(* IEC 61131-3 sources: volt/packages/volt-lsp-iec/test-corpus/pro2193/Device/Plc Logic/Application/09 Misc/Library Manager/L_TT1P_TechnologyModules (part 6) *)

(* ---- L_TT1P_WINDERTENSIONCTRLHIGH.pou ---- *)
FUNCTION_BLOCK L_TT1P_WINDERTENSIONCTRLHIGH EXTENDS TM_Winder
VAR_INPUT
	XENABLEINTERNALCONTROL : BOOL;
	XENABLE : BOOL;
	SCCTRLABC : scCtrl_ABC;
	XRESETERROR : BOOL;
	XREGULATORON : BOOL;
	XSTOP : BOOL;
	XHALT : BOOL;
	SCPAR : L_TT1P_scPar_WinderTensionCtrlHigh;
	MATERIALCOUNTERAXIS : L_MC1P_IAXIS_REF_POOL;
	SCACCESSPOINTS : L_TT1P_scAP_WinderTensionCtrlHigh;
	XMATERIALFEEDING : BOOL;
	XWINDINGDIRECTION : BOOL;
	XWINDINGDIRECTIONSTANDSTILL : BOOL;
	XLOADDIAM : BOOL;
	LRSETDIAM : LREAL;
	XHOLDDIAM : BOOL;
	XDIAMCALCREDUCED : BOOL;
	XSETMATERIALCOUNTER : BOOL;
	XWEBBREAKMONIT : BOOL;
	XJOGLINEPOS : BOOL;
	XJOGLINENEG : BOOL;
	XTRIMLINEPOS : BOOL;
	XTRIMLINENEG : BOOL;
	XSYNCLINEVEL : BOOL;
	XTENSCURVE : BOOL;
	LRSETTENS : LREAL;
	LRSETLINEVEL : LREAL;
	XTENSCTRL : BOOL;
	XFRICCMPS : BOOL;
	XACCCMPS : BOOL;
	LRMINERTIAADAPT : LREAL;
	LRACTTENSIN : LREAL;
	LRSETFRICADAPT : LREAL;
	LRTENSCTRLINFLUENCE : LREAL;
	XRESETPICTRL : BOOL;
	XRESETICTRL : BOOL;
	XEXECUTEIDENTFRIC : BOOL;
	XEXECUTEIDENTMINERTIA : BOOL;
	XADAPTSPDCTRLGAIN : BOOL;
	LRADAPTSPDCTRLGAINFACTOR : LREAL := 1;
END_VAR
VAR_OUTPUT
	XINTERNALCONTROLACTIVE : BOOL;
	ETMSTATE : L_TT1P_States;
	SCSTATUSABC : scStatus_ABC;
	XERROR : BOOL;
	XWARNING : BOOL;
	EERRORID : L_IE1P_Error;
	SCERRORINFO : L_TT1P_scErrorInfo;
	XAXISENABLED : BOOL;
	SCSIGNALFLOW : L_TT1P_scSF_WinderTensionCtrlHigh;
	XDONE : BOOL;
	XBUSY : BOOL;
	XSYNCHRONISED : BOOL;
	XACCDECSYNC : BOOL;
	XUNWIND : BOOL;
	XWEBBREAK : BOOL;
	XHOLDDIAMACTIVE : BOOL;
	XDIAMMAX : BOOL;
	XDIAMMIN : BOOL;
	LRSETDIAMOUT : LREAL;
	LRSETDIAMSCALEDOUT : LREAL;
	LRMATERIALCOUNTER : LREAL;
	LRSETLINEVELSCALEDOUT : LREAL;
	LRACTTOTALTRQSCALED : LREAL;
	LRWNDSPDREF : LREAL;
	XWNDSPDLIMIT : BOOL;
	LRLIMITLINEVEL : LREAL;
	LRSETMINERTIAOUT : LREAL;
	LRSETTENSSCALEDOUT : LREAL;
	LRSETTENSTRQSCALEDOUT : LREAL;
	LRSETFRICTRQSCALEDOUT : LREAL;
	LRSETACCTRQSCALEDOUT : LREAL;
	LRACTTENSSCALED : LREAL;
	LRSETTENSCTRLSCALEDOUT : LREAL;
	LRIDENTMINERTIA : LREAL;
	LRSETSPDCTRLGAINADAPTOUT : LREAL;
END_VAR
VAR_IN_OUT
	AXIS : AXIS_REF;
	PERSISTENTVAR : L_TT1P_PersistentVarWinder;
	ALRFRICTIONCURVE1 : ARRAY [1..66] OF LREAL;
	ALRFRICTIONCURVE2 : ARRAY [1..66] OF LREAL;
	ALRFRICTIONCURVE3 : ARRAY [1..66] OF LREAL;
	ALRFRICTIONCURVE4 : ARRAY [1..66] OF LREAL;
END_VAR
VAR
	TM_INT : _TM_WinderTensionCtrlHigh;
	PPAR : POINTER TO L_TT1P_scPar_WinderTensionCtrlHigh;
	PPAR_INT : POINTER TO L_TT1P_scPar_WinderTensionCtrlHigh;
	XISHOMED : BOOL;
	XHOMEEXECUTE : BOOL;
	XHOMEABSSWITCH : BOOL;
	XJOGPOS : BOOL;
	XJOGNEG : BOOL;
END_VAR
END_FUNCTION_BLOCK

METHOD CALL_COUPLINGREELSPEEDLIMIT
END_METHOD

METHOD CALL_DECOUPLINGREELSPEEDLIMIT
END_METHOD

METHOD GET_ESTATE : L_TT1P_States
END_METHOD

METHOD GET_ETMSTATE : L_TT1P_States
END_METHOD

METHOD GET_LRACTACCTRQ : LREAL
END_METHOD

METHOD GET_LRACTFRICTRQ : LREAL
END_METHOD

METHOD GET_LRACTMOTORTORQUE : LREAL
END_METHOD

METHOD GET_LRACTTENSTRQ : LREAL
END_METHOD

METHOD GET_LRCALCDIAMDIST : LREAL
END_METHOD

METHOD GET_LRCALCDIAMLINESPEED : LREAL
END_METHOD

METHOD GET_LRCALCDIAMREELSPEED : LREAL
END_METHOD

METHOD GET_LRFEEDCONSTANT : LREAL
END_METHOD

METHOD GET_LRLOWERSPEEDLIMIT : LREAL
END_METHOD

METHOD GET_LRMOTORTORQUEREF : LREAL
END_METHOD

METHOD GET_LRRAMPGENOUT : LREAL
END_METHOD

METHOD GET_LRREELSPEEDREF : LREAL
END_METHOD

METHOD GET_LRSETMOTORTORQUE : LREAL
END_METHOD

METHOD GET_LRSETSPEEDCTRLGAINADAPT : LREAL
END_METHOD

METHOD GET_LRSETTOTALTORQUE : LREAL
END_METHOD

METHOD GET_LRSPEEDLOWERLIMIT : LREAL
END_METHOD

METHOD GET_LRSPEEDUPPERLIMIT : LREAL
END_METHOD

METHOD GET_LRTASKCYCLE : LREAL
END_METHOD

METHOD GET_LRTENSCTRLOUT : LREAL
END_METHOD

METHOD GET_LRTENSCURVEOUT : LREAL
END_METHOD

METHOD GET_LRUPPERSPEEDLIMIT : LREAL
END_METHOD

METHOD GET_LRVARMINERTIASCALED : LREAL
END_METHOD

METHOD GET_LRWINDERTORQUEREF : LREAL
END_METHOD

METHOD GET_XCOMMUNICATION : BOOL
END_METHOD

METHOD GET_XDIAMWEBBREAKENABLE : BOOL
VAR_OUTPUT
	XUNIDIRECT : BOOL;
	XUNWINDACTIVE : BOOL;
END_VAR
END_METHOD

METHOD RESET_SYSTEMFAULT
END_METHOD

METHOD SET_SYSTEMFAULT
VAR_INPUT
	IN : L_IE1P_Error;
END_VAR
END_METHOD

METHOD SET_ALRPROCESSCTRLXVALUES
VAR_INPUT
	ALRPROCESSCTRLXVALUES : ARRAY [1..5] OF LREAL := [5(0)];
END_VAR
END_METHOD

METHOD SET_ALRPROCESSCTRLYVALUES
VAR_INPUT
	ALRPROCESSCTRLYVALUES : ARRAY [1..5] OF LREAL := [1, 4(0)];
END_VAR
END_METHOD

METHOD SET_ESTATE
VAR_INPUT
	IN : L_TT1P_States;
END_VAR
END_METHOD

METHOD SET_LRFEEDCONSTANT
VAR_INPUT
	LRIN : LREAL := 0;
END_VAR
END_METHOD

METHOD SET_LRPICTRLINTVALUE
VAR_INPUT
	LRIN : LREAL := 0;
END_VAR
END_METHOD

METHOD SET_LRPROCESSCTRLACC
VAR_INPUT
	LRPROCESSCTRLACC : LREAL := 0.0;
END_VAR
END_METHOD

METHOD SET_LRPROCESSCTRLDEC
VAR_INPUT
	LRPROCESSCTRLDEC : LREAL := 0.0;
END_VAR
END_METHOD

METHOD SET_LRPROCESSCTRLGAINADAPT
VAR_INPUT
	LRPROCESSCTRLGAINADAPT : LREAL := 1;
END_VAR
END_METHOD

METHOD SET_LRPROCESSCTRLINTVALUE
VAR_INPUT
	LRPROCESSCTRLINTVALUE : LREAL := 0.0;
END_VAR
END_METHOD

METHOD SET_LRPROCESSCTRLREDGAIN
VAR_INPUT
	LRPROCESSCTRLREDGAIN : LREAL := 0.0;
END_VAR
END_METHOD

METHOD SET_LRPROCESSCTRLREDRANGE
VAR_INPUT
	LRPROCESSCTRLREDRANGE : LREAL := 0.0;
END_VAR
END_METHOD

METHOD SET_LRREFERENCEMOTORTORQUE
VAR_INPUT
	LRIN : LREAL := 0;
END_VAR
END_METHOD

METHOD SET_LRREFERENCEREELSPEED
VAR_INPUT
	LRIN : LREAL := 0;
END_VAR
END_METHOD

METHOD SET_LRSPEEDOFFSET
VAR_INPUT
	LRIN : LREAL := 0;
END_VAR
END_METHOD

METHOD SET_LRTORQUEOFFSET
VAR_INPUT
	LRIN : LREAL := 0;
END_VAR
END_METHOD

METHOD SET_RPROCESSCTRLDELAYTIME
VAR_INPUT
	RPROCESSCTRLDELAYTIME : REAL := 0.0;
END_VAR
END_METHOD

METHOD SET_RPROCESSCTRLRATEDTIME
VAR_INPUT
	RPROCESSCTRLRATEDTIME : REAL := 0.0;
END_VAR
END_METHOD

METHOD SET_XPICTRLLOADINTVALUE
VAR_INPUT
	XIN : BOOL := FALSE;
END_VAR
END_METHOD

METHOD SET_XPROCESSCTRLLOADINTVALUE
VAR_INPUT
	XPROCESSCTRLLOADINTVALUE : BOOL := FALSE;
END_VAR
END_METHOD

METHOD SET_XSPEEDLIMITENABLEDEXT
VAR_INPUT
	XIN : BOOL := TRUE;
END_VAR
END_METHOD

METHOD SET_XWEBBREAK
VAR_INPUT
	XIN : BOOL := FALSE;
END_VAR
END_METHOD

(* ---- L_TT1P_WINDERTENSIONCTRLSTATE.pou ---- *)
FUNCTION_BLOCK L_TT1P_WINDERTENSIONCTRLSTATE EXTENDS TM_Winder
VAR_INPUT
	XENABLEINTERNALCONTROL : BOOL;
	XENABLE : BOOL;
	SCCTRLABC : scCtrl_ABC;
	XRESETERROR : BOOL;
	XREGULATORON : BOOL;
	XSTOP : BOOL;
	XHALT : BOOL;
	SCPAR : L_TT1P_scPar_WinderTensionCtrlState;
	MATERIALCOUNTERAXIS : L_MC1P_IAXIS_REF_POOL;
	SCACCESSPOINTS : L_TT1P_scAP_WinderTensionCtrlState;
	XMATERIALFEEDING : BOOL;
	XWINDINGDIRECTION : BOOL;
	XWINDINGDIRECTIONSTANDSTILL : BOOL;
	XLOADDIAM : BOOL;
	LRSETDIAM : LREAL;
	XHOLDDIAM : BOOL;
	XDIAMCALCREDUCED : BOOL;
	XSETMATERIALCOUNTER : BOOL;
	XWEBBREAKMONIT : BOOL;
	XJOGLINEPOS : BOOL;
	XJOGLINENEG : BOOL;
	XTRIMLINEPOS : BOOL;
	XTRIMLINENEG : BOOL;
	XSYNCLINEVEL : BOOL;
	XTENSCURVE : BOOL;
	LRSETTENS : LREAL;
	LRSETLINEVEL : LREAL;
	XTENSCTRL : BOOL;
	XFRICCMPS : BOOL;
	XACCCMPS : BOOL;
	LRMINERTIAADAPT : LREAL := 1;
	LRACTTENSIN : LREAL;
	LRSETFRICADAPT : LREAL;
	LRTENSCTRLINFLUENCE : LREAL;
	XRESETPICTRL : BOOL;
	XRESETICTRL : BOOL;
	XEXECUTEIDENTFRIC : BOOL;
END_VAR
VAR_OUTPUT
	XINTERNALCONTROLACTIVE : BOOL;
	ETMSTATE : L_TT1P_States;
	SCSTATUSABC : scStatus_ABC;
	XERROR : BOOL;
	XWARNING : BOOL;
	EERRORID : L_IE1P_Error;
	SCERRORINFO : L_TT1P_scErrorInfo;
	XAXISENABLED : BOOL;
	SCSIGNALFLOW : L_TT1P_scSF_WinderTensionCtrlState;
	XDONE : BOOL;
	XBUSY : BOOL;
	XSYNCHRONISED : BOOL;
	XACCDECSYNC : BOOL;
	XUNWIND : BOOL;
	XWEBBREAK : BOOL;
	XHOLDDIAMACTIVE : BOOL;
	XDIAMMAX : BOOL;
	XDIAMMIN : BOOL;
	LRSETDIAMOUT : LREAL;
	LRSETDIAMSCALEDOUT : LREAL;
	LRMATERIALCOUNTER : LREAL;
	LRSETLINEVELSCALEDOUT : LREAL;
	LRACTTOTALTRQSCALED : LREAL;
	LRWNDSPDREF : LREAL;
	XWNDSPDLIMIT : BOOL;
	LRLIMITLINEVEL : LREAL;
	LRSETMINERTIAOUT : LREAL;
	LRSETTENSSCALEDOUT : LREAL;
	LRSETTENSTRQSCALEDOUT : LREAL;
	LRSETFRICTRQSCALEDOUT : LREAL;
	LRSETACCTRQSCALEDOUT : LREAL;
	LRACTTENSSCALED : LREAL;
	LRSETTENSCTRLSCALEDOUT : LREAL;
END_VAR
VAR_IN_OUT
	AXIS : AXIS_REF;
	PERSISTENTVAR : L_TT1P_PersistentVarWinder;
	ALRFRICTIONCURVE1 : ARRAY [1..66] OF LREAL;
	ALRFRICTIONCURVE2 : ARRAY [1..66] OF LREAL;
	ALRFRICTIONCURVE3 : ARRAY [1..66] OF LREAL;
	ALRFRICTIONCURVE4 : ARRAY [1..66] OF LREAL;
END_VAR
VAR
	TM_INT : _TM_WinderTensionCtrlState;
	PPAR : POINTER TO L_TT1P_scPar_WinderTensionCtrlState;
	PPAR_INT : POINTER TO L_TT1P_scPar_WinderTensionCtrlState;
	XISHOMED : BOOL;
	XHOMEEXECUTE : BOOL;
	XHOMEABSSWITCH : BOOL;
	XJOGPOS : BOOL;
	XJOGNEG : BOOL;
END_VAR
END_FUNCTION_BLOCK

METHOD CALL_COUPLINGREELSPEEDLIMIT
END_METHOD

METHOD CALL_DECOUPLINGREELSPEEDLIMIT
END_METHOD

METHOD GET_ESTATE : L_TT1P_States
END_METHOD

METHOD GET_ETMSTATE : L_TT1P_States
END_METHOD

METHOD GET_LRACTACCTRQ : LREAL
END_METHOD

METHOD GET_LRACTFRICTRQ : LREAL
END_METHOD

METHOD GET_LRACTMOTORTORQUE : LREAL
END_METHOD

METHOD GET_LRACTTENSTRQ : LREAL
END_METHOD

METHOD GET_LRCALCDIAMDIST : LREAL
END_METHOD

METHOD GET_LRCALCDIAMLINESPEED : LREAL
END_METHOD

METHOD GET_LRCALCDIAMREELSPEED : LREAL
END_METHOD

METHOD GET_LRFEEDCONSTANT : LREAL
END_METHOD

METHOD GET_LRLOWERSPEEDLIMIT : LREAL
END_METHOD

METHOD GET_LRMOTORTORQUEREF : LREAL
END_METHOD

METHOD GET_LRRAMPGENOUT : LREAL
END_METHOD

METHOD GET_LRREELSPEEDREF : LREAL
END_METHOD

METHOD GET_LRSETMOTORTORQUE : LREAL
END_METHOD

METHOD GET_LRSETSPEEDCTRLGAINADAPT : LREAL
END_METHOD

METHOD GET_LRSETTOTALTORQUE : LREAL
END_METHOD

METHOD GET_LRSPEEDLOWERLIMIT : LREAL
END_METHOD

METHOD GET_LRSPEEDUPPERLIMIT : LREAL
END_METHOD

METHOD GET_LRTASKCYCLE : LREAL
END_METHOD

METHOD GET_LRTENSCTRLOUT : LREAL
END_METHOD

METHOD GET_LRTENSCURVEOUT : LREAL
END_METHOD

METHOD GET_LRUPPERSPEEDLIMIT : LREAL
END_METHOD

METHOD GET_LRVARMINERTIASCALED : LREAL
END_METHOD

METHOD GET_LRWINDERTORQUEREF : LREAL
END_METHOD

METHOD GET_XCOMMUNICATION : BOOL
END_METHOD

METHOD GET_XDIAMWEBBREAKENABLE : BOOL
VAR_OUTPUT
	XUNIDIRECT : BOOL;
	XUNWINDACTIVE : BOOL;
END_VAR
END_METHOD

METHOD RESET_SYSTEMFAULT
END_METHOD

METHOD SET_SYSTEMFAULT
VAR_INPUT
	IN : L_IE1P_Error;
END_VAR
END_METHOD

METHOD SET_ALRPROCESSCTRLXVALUES
VAR_INPUT
	ALRPROCESSCTRLXVALUES : ARRAY [1..5] OF LREAL := [5(0)];
END_VAR
END_METHOD

METHOD SET_ALRPROCESSCTRLYVALUES
VAR_INPUT
	ALRPROCESSCTRLYVALUES : ARRAY [1..5] OF LREAL := [1, 4(0)];
END_VAR
END_METHOD

METHOD SET_ESTATE
VAR_INPUT
	IN : L_TT1P_States;
END_VAR
END_METHOD

METHOD SET_LRFEEDCONSTANT
VAR_INPUT
	LRIN : LREAL := 0;
END_VAR
END_METHOD

METHOD SET_LRPICTRLINTVALUE
VAR_INPUT
	LRIN : LREAL := 0;
END_VAR
END_METHOD

METHOD SET_LRPROCESSCTRLACC
VAR_INPUT
	LRPROCESSCTRLACC : LREAL := 0.0;
END_VAR
END_METHOD

METHOD SET_LRPROCESSCTRLDEC
VAR_INPUT
	LRPROCESSCTRLDEC : LREAL := 0.0;
END_VAR
END_METHOD

METHOD SET_LRPROCESSCTRLGAINADAPT
VAR_INPUT
	LRPROCESSCTRLGAINADAPT : LREAL := 1;
END_VAR
END_METHOD

METHOD SET_LRPROCESSCTRLINTVALUE
VAR_INPUT
	LRPROCESSCTRLINTVALUE : LREAL := 0.0;
END_VAR
END_METHOD

METHOD SET_LRPROCESSCTRLREDGAIN
VAR_INPUT
	LRPROCESSCTRLREDGAIN : LREAL := 0.0;
END_VAR
END_METHOD

METHOD SET_LRPROCESSCTRLREDRANGE
VAR_INPUT
	LRPROCESSCTRLREDRANGE : LREAL := 0.0;
END_VAR
END_METHOD

METHOD SET_LRREFERENCEMOTORTORQUE
VAR_INPUT
	LRIN : LREAL := 0;
END_VAR
END_METHOD

METHOD SET_LRREFERENCEREELSPEED
VAR_INPUT
	LRIN : LREAL := 0;
END_VAR
END_METHOD

METHOD SET_LRSPEEDOFFSET
VAR_INPUT
	LRIN : LREAL := 0;
END_VAR
END_METHOD

METHOD SET_LRTORQUEOFFSET
VAR_INPUT
	LRIN : LREAL := 0;
END_VAR
END_METHOD

METHOD SET_RPROCESSCTRLDELAYTIME
VAR_INPUT
	RPROCESSCTRLDELAYTIME : REAL := 0.0;
END_VAR
END_METHOD

METHOD SET_RPROCESSCTRLRATEDTIME
VAR_INPUT
	RPROCESSCTRLRATEDTIME : REAL := 0.0;
END_VAR
END_METHOD

METHOD SET_XPICTRLLOADINTVALUE
VAR_INPUT
	XIN : BOOL := FALSE;
END_VAR
END_METHOD

METHOD SET_XPROCESSCTRLLOADINTVALUE
VAR_INPUT
	XPROCESSCTRLLOADINTVALUE : BOOL := FALSE;
END_VAR
END_METHOD

METHOD SET_XSPEEDLIMITENABLEDEXT
VAR_INPUT
	XIN : BOOL := TRUE;
END_VAR
END_METHOD

METHOD SET_XWEBBREAK
VAR_INPUT
	XIN : BOOL := FALSE;
END_VAR
END_METHOD

(* ---- TM_WINDER.pou ---- *)
FUNCTION_BLOCK TM_WINDER
END_FUNCTION_BLOCK

METHOD CALL_SMC_READPARAMETEREXT
VAR_INPUT
	XENABLE : BOOL;
	WCODENUMBER : WORD;
	BYSUBCODE : BYTE;
END_VAR
VAR_OUTPUT
	XVALID : BOOL;
	XBUSY : BOOL;
	XERROR : BOOL;
	WERRORID : WORD;
	DWVALUE : DWORD;
END_VAR
END_METHOD

METHOD CALL_WRITEPARAMETEREXT
VAR_INPUT
	XEXECUTE : BOOL;
	WCODENUMBER : WORD;
	BYSUBCODE : BYTE;
	BYLENGTH : BYTE;
	DNVALUE : DINT;
END_VAR
VAR_OUTPUT
	XDONE : BOOL;
	XBUSY : BOOL;
	XERROR : BOOL;
	WERRORID : WORD;
END_VAR
END_METHOD

METHOD CALL_WRITEPARAMETEREXT2
VAR_INPUT
	XEXECUTE : BOOL;
	WCODENUMBER : WORD;
	BYSUBCODE : BYTE;
	BYLENGTH : BYTE;
	DNVALUE : DINT;
END_VAR
VAR_OUTPUT
	XDONE : BOOL;
	XBUSY : BOOL;
	XERROR : BOOL;
	WERRORID : WORD;
END_VAR
END_METHOD

METHOD GET_ESTATE : L_TT1P_States
END_METHOD

METHOD GET_ETMSTATE : L_TT1P_States
END_METHOD

METHOD GET_FSCALEFACTOR : LREAL
END_METHOD

METHOD GET_LRACTMOTORTORQUE : LREAL
END_METHOD

METHOD GET_LRCALCDIAMDIST : LREAL
END_METHOD

METHOD GET_LRFEEDCONSTANT : LREAL
END_METHOD

METHOD GET_LRLOWERSPEEDLIMIT : LREAL
END_METHOD

METHOD GET_LRMOTORTORQUEREF : LREAL
END_METHOD

METHOD GET_LRREELSPEEDREF : LREAL
END_METHOD

METHOD GET_LRSETMOTORTORQUE : LREAL
END_METHOD

METHOD GET_LRSETSPEEDCTRLGAINADAPT : LREAL
END_METHOD

METHOD GET_LRSETTOTALTORQUE : LREAL
END_METHOD

METHOD GET_LRTASKCYCLE : LREAL
END_METHOD

METHOD GET_LRUPPERSPEEDLIMIT : LREAL
END_METHOD

METHOD GET_LRVARMINERTIASCALED : LREAL
END_METHOD

METHOD GET_LRWINDERTORQUEREF : LREAL
END_METHOD

METHOD GET_WCHECKAXISTYP : WORD
END_METHOD

METHOD GET_XCOMMUNICATION : BOOL
END_METHOD

METHOD GET_XDIAMWEBBREAKENABLE : BOOL
VAR_OUTPUT
	XUNIDIRECT : BOOL;
	XUNWINDACTIVE : BOOL;
END_VAR
END_METHOD

METHOD RESET_SYSTEMFAULT
END_METHOD

METHOD SET_SYSTEMFAULT
VAR_INPUT
	IN : L_IE1P_Error;
END_VAR
END_METHOD

METHOD SET_WNDAXISEXTENSION_READY
END_METHOD

METHOD SET_ESTATE
VAR_INPUT
	IN : L_TT1P_States;
END_VAR
END_METHOD

METHOD SET_LRFEEDCONSTANT
VAR_INPUT
	LRIN : LREAL := 0;
END_VAR
END_METHOD

METHOD SET_LRREFERENCEMOTORTORQUE
VAR_INPUT
	LRIN : LREAL := 0;
END_VAR
END_METHOD

METHOD SET_LRREFERENCEREELSPEED
VAR_INPUT
	LRIN : LREAL := 0;
END_VAR
END_METHOD

METHOD SET_LRSPEEDOFFSET
VAR_INPUT
	LRIN : LREAL := 0;
END_VAR
END_METHOD

METHOD SET_LRTORQUEOFFSET
VAR_INPUT
	LRIN : LREAL := 0;
END_VAR
END_METHOD

METHOD SET_XSPEEDLIMITENABLEDEXT
VAR_INPUT
	XIN : BOOL := TRUE;
END_VAR
END_METHOD

METHOD SET_XWEBBREAK
VAR_INPUT
	XIN : BOOL := FALSE;
END_VAR
END_METHOD
